{attribute 'qualified_only'}
VAR_GLOBAL
	//DEVICES
	VTD:  VTD_Control_DUT;
	ECnv:  ECnv_Control_DUT;
	LCnv:  ARRAY[1..6] OF Buffer_Cnv_Control_DUT;
	Turn_Table: Turn_Table_Control_DUT;
	TBCnv:  TBCnv_Control_DUT;
	Pop_Up_Cnv: ARRAY[1..2] OF PopUp_Control_DUT;
	Roller_Cnv: ARRAY[1..5] OF Roller_Control_DUT;
	Chain_Cnv: Chain_Control_DUT;
	VTDBarcode_Station:  ARRAY[1..3] OF Barcode_Station_DUT;
	Profiling_Station: ARRAY[1..2] OF Profiling_Station_DUT;
	
	//ORDER TABLES COMMANDS
	VTD_Order_Table:  WMS_OPC_UA_DUT;
	Carousel_Order_Table:  WMS_OPC_UA_DUT;
	
	Shuttles_Position:  ARRAY[1..10] OF Shuttle_Position_UDT;
	
	Gate_Station:  ARRAY[1..2] OF Gate_Station_DUT;
	Charger_Level:  ARRAY[1..6] OF Charger_DUT;
END_VAR

(* stored: Version 1.1.0.1
   GVL Control: Id {5e6952d4-e20c-4a7f-aad7-0649e4f09d9f} *)
